// TIA Portal V21 export
FUNCTION_BLOCK "FB_StarterScl"   // FB104, SCL
TITLE = Пускатель насоса (SCL)
{ S7_Optimized_Access := 'TRUE' }
AUTHOR : WTP2
FAMILY : Drives
VERSION : 0.1
// Пускатель насоса с контролем обратной связи (один блок на LAD, FBD, STL, SCL).
// 1. Пуск/стоп — SR с битом-операндом xRunMem: S = xStart AND xInterlock; R1 = xStop OR NOT xInterlock OR xFault.
//    SR S7: сначала S, затем R1 — при S = R1 = 1 (Пуск и Стоп одновременно) бит сброшен. xRun := xRunMem.
// 2. Контроль обратной связи: TON tonFeedback (IN = xRun AND NOT xFeedback, PT = tFeedbackTime).
// 3. Авария с самоподхватом: xFault := (tonFeedback.Q OR xFault) AND NOT xReset.
// 4. Счётчик пусков: по фронту xRun (бит памяти xEdgeMem) iStarts := iStarts + 1.
// Порядок сетей 1-4; xFault в сети 1 — значение прошлого вызова.
// stored: AutoNumber false, SetENOAutomatically false
   VAR_INPUT
      xStart : Bool;   // Пуск (кнопка)
      xStop : Bool;   // Стоп (кнопка, TRUE — нажата)
      xInterlock : Bool := TRUE;   // Блокировки в норме, пуск разрешён
      xFeedback : Bool;   // Обратная связь контактора
      tFeedbackTime : Time := T#2S;   // Допустимое время без обратной связи
      xReset : Bool;   // Сброс аварии
   END_VAR
   VAR_OUTPUT
      xRun : Bool;   // Команда контактору
      xFault : Bool;   // Авария: нет обратной связи
      iStarts : Int;   // Число пусков
   END_VAR
   VAR
      xRunMem : Bool;   // Бит-операнд SR пуска
      xEdgeMem : Bool;   // Бит памяти фронта xRun
      tonFeedback : TON_TIME;   // Таймер контроля обратной связи
   END_VAR
BEGIN
// Пускатель
// Логика пускателя целиком
   // 1. SR с битом xRunMem: сначала S, затем R1 (сброс главнее)
   IF #xStart AND #xInterlock THEN
       #xRunMem := TRUE;
   END_IF;
   IF #xStop OR NOT #xInterlock OR #xFault THEN
       #xRunMem := FALSE;
   END_IF;
   #xRun := #xRunMem;
   // 2. Контроль обратной связи
   #tonFeedback(IN := #xRun AND NOT #xFeedback, PT := #tFeedbackTime);
   // 3. Авария с самоподхватом
   #xFault := (#tonFeedback.Q OR #xFault) AND NOT #xReset;
   // 4. Счётчик пусков по фронту xRun
   IF #xRun AND NOT #xEdgeMem THEN
       #iStarts := #iStarts + 1;
   END_IF;
   #xEdgeMem := #xRun;
END_FUNCTION_BLOCK
